Fanuc KAREL source: KO00013.KL

PROGRAM KO00013
%NOLOCKGROUP
VAR
  P1: XYZWPR
  P2: XYZWPR
  P3: XYZWPR
  P4: XYZWPR
  OUT: POSITION
BEGIN
  OUT = FRAME(P1, P2, P3, P4)
END KO00013
